(* Logix 5000 project; controller NWGG_Treater_Dayton vendor 1 type 14 code 238 rev 35.11; software revision 35.00 *)
// Treater at the Walla Walla Seed Plant

TASK MainTask (continuous, watchdog 500 ms) : MainProgram, Pumps, ColorBlending
TASK SafetyTask (periodic, rate 20 ms, priority 10, watchdog 20 ms, safety) : SafetyProgram

MODULES
   Local : vendor 1 type 14 code 238 (5069 0, rev 35.11)
      Pump_8 : PowerFlex 525-EENET (Ethernet 192.168.1.64, rev 7.1, Output RPI 20 ms)
      Pump_9 : PowerFlex 525-EENET (Ethernet 192.168.1.65, rev 7.1, Output RPI 20 ms)
      Pump_19 : PowerFlex 525-EENET (Ethernet 192.168.1.75, rev 7.1, Output RPI 20 ms)
      Pump_10 : PowerFlex 525-EENET (Ethernet 192.168.1.66, rev 7.1, Output RPI 20 ms)
      Pump_18 : PowerFlex 525-EENET (Ethernet 192.168.1.74, rev 7.1, Output RPI 20 ms)
      Pump_16 : PowerFlex 525-EENET (Ethernet 192.168.1.72, rev 7.1, Output RPI 20 ms)
      Pump_3 : PowerFlex 525-EENET (Ethernet 192.168.1.59, rev 7.1, Output RPI 20 ms)
      Treater_Drive : PowerFlex 525-EENET (Ethernet 192.168.1.81, rev 7.1, Output RPI 20 ms)
      Pump_21 : PowerFlex 525-EENET (Ethernet 192.168.1.77, rev 7.1, Output RPI 20 ms)
      Pump_6 : PowerFlex 525-EENET (Ethernet 192.168.1.62, rev 7.1, Output RPI 20 ms)
      Pump_20 : PowerFlex 525-EENET (Ethernet 192.168.1.76, rev 7.1, Output RPI 20 ms)
      Pump_22 : PowerFlex 525-EENET (Ethernet 192.168.1.78, rev 7.1, Output RPI 20 ms)
      Pump_14 : PowerFlex 525-EENET (Ethernet 192.168.1.70, rev 7.1, Output RPI 20 ms)
      Pump_13 : PowerFlex 525-EENET (Ethernet 192.168.1.69, rev 7.1, Output RPI 20 ms)
      Pump_15 : PowerFlex 525-EENET (Ethernet 192.168.1.71, rev 7.1, Output RPI 20 ms)
      Pump_7 : PowerFlex 525-EENET (Ethernet 192.168.1.63, rev 7.1, Output RPI 20 ms)
      Pump_5 : PowerFlex 525-EENET (Ethernet 192.168.1.61, rev 7.1, Output RPI 20 ms)
      Pump_12 : PowerFlex 525-EENET (Ethernet 192.168.1.68, rev 7.1, Output RPI 20 ms)
      Pump_2 : PowerFlex 525-EENET (Ethernet 192.168.1.58, rev 7.1, Output RPI 20 ms)
      Pump_1 : PowerFlex 525-EENET (Ethernet 192.168.1.57, rev 7.1, Output RPI 20 ms)
      Pump_11 : PowerFlex 525-EENET (Ethernet 192.168.1.67, rev 7.1, Output RPI 20 ms)
      Pump_17 : PowerFlex 525-EENET (Ethernet 192.168.1.73, rev 7.1, Output RPI 20 ms)
      Pump_4 : PowerFlex 525-EENET (Ethernet 192.168.1.60, rev 7.1, Output RPI 20 ms)
      Flex_IO_Adapter : 1794-AENTR (Ethernet 192.168.1.100, rev 1.1, Output RPI 20 ms)
         AC_Input : 1794-IA16 (Flex 2, rev 1.1)
         AC_Output : vendor 1 type 7 code 48 (Flex 3, rev 1.1)
         Analog_In_1 : vendor 1 type 10 code 25 (Flex 0, rev 2.1, Input RPI 80 ms)
         Analog_In_2 : vendor 1 type 10 code 25 (Flex 1, rev 2.1, Input RPI 80 ms)
      Scale_13 : vendor 666 type 12 code 16898 (Ethernet 192.168.1.123, rev 1.1, StandardDataDriven RPI 2 ms)
      Scale_22 : vendor 666 type 12 code 16898 (Ethernet 192.168.1.132, rev 1.1, StandardDataDriven RPI 2 ms)   // Pea Slurry
      Scale_9 : vendor 666 type 12 code 16898 (Ethernet 192.168.1.119, rev 1.1, StandardDataDriven RPI 2 ms)
      Scale_17 : vendor 666 type 12 code 16898 (Ethernet 192.168.1.127, rev 1.1, StandardDataDriven RPI 2 ms)
      Scale_8 : vendor 666 type 12 code 16898 (Ethernet 192.168.1.118, rev 1.1, StandardDataDriven RPI 2 ms)
      Scale_20 : vendor 666 type 12 code 16898 (Ethernet 192.168.1.130, rev 1.1, StandardDataDriven RPI 2 ms)
      Scale_19 : vendor 666 type 12 code 16898 (Ethernet 192.168.1.129, rev 1.1, StandardDataDriven RPI 2 ms)
      Scale_14 : vendor 666 type 12 code 16898 (Ethernet 192.168.1.124, rev 1.1, StandardDataDriven RPI 2 ms)
      Scale_6 : vendor 666 type 12 code 16898 (Ethernet 192.168.1.116, rev 1.1, StandardDataDriven RPI 2 ms)
      Scale_11 : vendor 666 type 12 code 16898 (Ethernet 192.168.1.121, rev 1.1, StandardDataDriven RPI 2 ms)
      Scale_21 : vendor 666 type 12 code 16898 (Ethernet 192.168.1.131, rev 1.1, StandardDataDriven RPI 2 ms)   // Small 3' By 3' Floor Scale
      Scale_1 : vendor 666 type 12 code 16898 (Ethernet 192.168.1.111, rev 1.1, StandardDataDriven RPI 2 ms)
      Scale_4 : vendor 666 type 12 code 16898 (Ethernet 192.168.1.114, rev 1.1, StandardDataDriven RPI 2 ms)
      Scale_18 : vendor 666 type 12 code 16898 (Ethernet 192.168.1.128, rev 1.1, StandardDataDriven RPI 2 ms)
      Scale_3 : vendor 666 type 12 code 16898 (Ethernet 192.168.1.113, rev 1.1, StandardDataDriven RPI 2 ms)
      Scale_5 : vendor 666 type 12 code 16898 (Ethernet 192.168.1.115, rev 1.1, StandardDataDriven RPI 2 ms)
      Scale_16 : vendor 666 type 12 code 16898 (Ethernet 192.168.1.126, rev 1.1, StandardDataDriven RPI 2 ms)
      Scale_2 : vendor 666 type 12 code 16898 (Ethernet 192.168.1.112, rev 1.1, StandardDataDriven RPI 2 ms)
      Scale_15 : vendor 666 type 12 code 16898 (Ethernet 192.168.1.125, rev 1.1, StandardDataDriven RPI 2 ms)
      Scale_10 : vendor 666 type 12 code 16898 (Ethernet 192.168.1.120, rev 1.1, StandardDataDriven RPI 2 ms)
      Scale_7 : vendor 666 type 12 code 16898 (Ethernet 192.168.1.117, rev 1.1, StandardDataDriven RPI 2 ms)
      Scale_12 : vendor 666 type 12 code 16898 (Ethernet 192.168.1.122, rev 1.1, StandardDataDriven RPI 2 ms)
      Water_Input : vendor 1 type 115 code 314 (5069 1, rev 2.1, StandardDataDriven RPI 100 ms)   // Input for Water Flow
END_MODULES

ADD_ON_INSTRUCTION Analog_Pump_Control   (* revision 1.0 *)
VAR_IN_OUT
   Pump_Drive_Out : AB:PowerFlex525V_EENET_Drive:O:0; {required}   // Pump Output
   Pump_Drive_In : AB:PowerFlex525V_EENET_Drive:I:0; {required}   // Pump Input
   Treater_Pump : Treater_Pump; {required}
        .Current_Oz_Rate   // This is the rate adjusted for the Current flow of grain reflected by the muiltliplier
END_VAR
VAR_INPUT
   Grain_Flow_CWT : REAL; {access None, required}
   Pump_Reversed : BOOL; {access Read Only, required}
END_VAR
VAR_IN_OUT
   Values : Analog_Gallon_Values; {required}   // Stored Values
   Analog_Raw_Counts : REAL; {required}
END_VAR
VAR_INPUT
   Start_Treating : BOOL; {access Read Only, required}
END_VAR
VAR
   Empty_String : STRING; {access None}
   PMC : Pump_Motor_Control; {access None}
   AnalogRate : Analog_Rate; {access None}
END_VAR

ROUTINE Logic   (* ladder *)
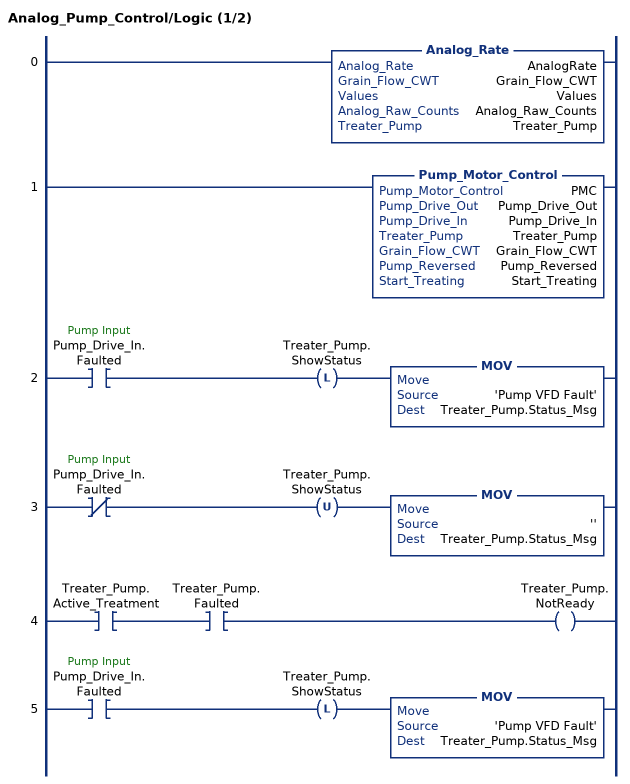
   0: Analog_Rate(AnalogRate,Grain_Flow_CWT,Values,Analog_Raw_Counts,Treater_Pump);
   1: Pump_Motor_Control(PMC,Pump_Drive_Out,Pump_Drive_In,Treater_Pump,Grain_Flow_CWT,Pump_Reversed,Start_Treating);
   2: XIC(Pump_Drive_In.Faulted)OTL(Treater_Pump.ShowStatus)MOV('Pump VFD Fault',Treater_Pump.Status_Msg);
   3: XIO(Pump_Drive_In.Faulted)OTU(Treater_Pump.ShowStatus)MOV('',Treater_Pump.Status_Msg);
   4: XIC(Treater_Pump.Active_Treatment)XIC(Treater_Pump.Faulted)OTE(Treater_Pump.NotReady);
   5: XIC(Pump_Drive_In.Faulted)OTL(Treater_Pump.ShowStatus)MOV('Pump VFD Fault',Treater_Pump.Status_Msg);
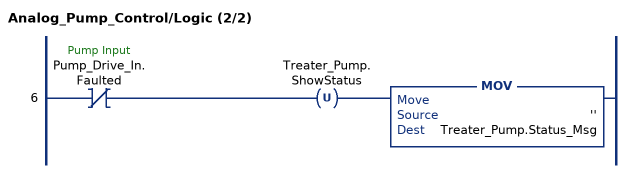
   6: XIO(Pump_Drive_In.Faulted)OTU(Treater_Pump.ShowStatus)MOV('',Treater_Pump.Status_Msg);
END_ROUTINE
END_ADD_ON_INSTRUCTION

ADD_ON_INSTRUCTION Analog_Rate   (* revision 1.0 *)
VAR_INPUT
   Grain_Flow_CWT : REAL; {access None, required}
END_VAR
VAR_IN_OUT
   Values : Analog_Gallon_Values; {required}   // Stored Values
END_VAR
VAR_INPUT
   Analog_Raw_Counts : REAL; {access Read Only, required}   // Values From CT
END_VAR
VAR_IN_OUT
   Treater_Pump : Treater_Pump; {required}
END_VAR

ROUTINE Logic   (* ladder *)
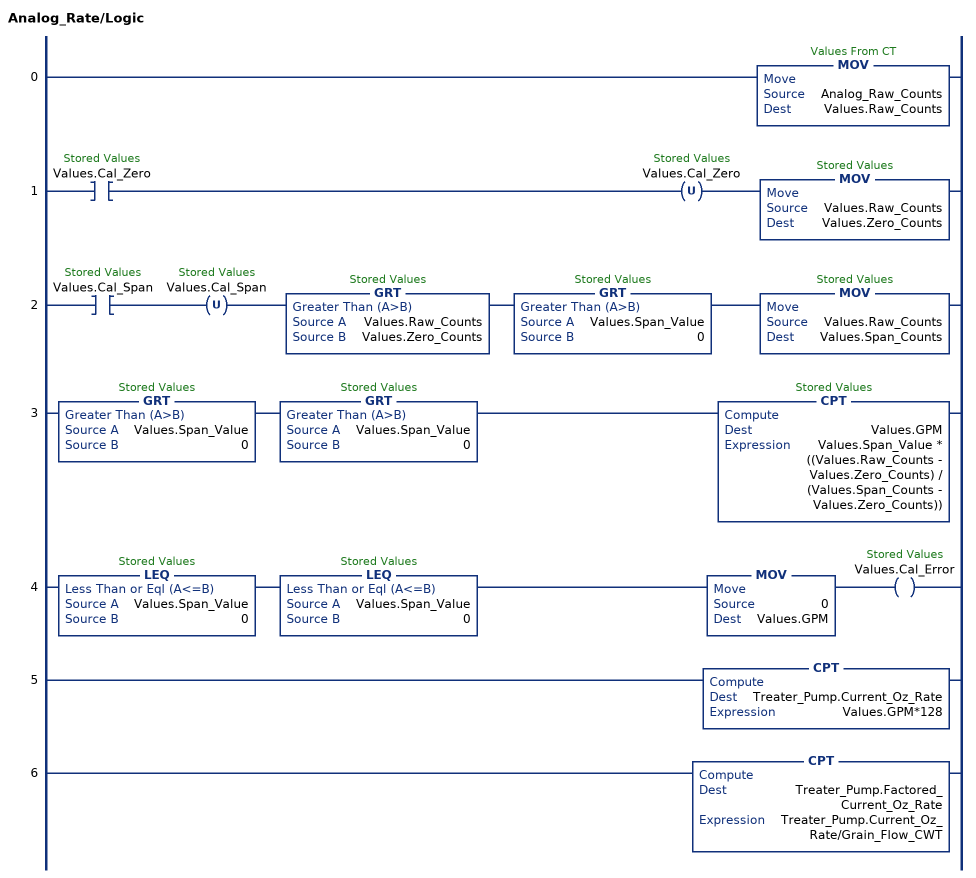
   0: MOV(Analog_Raw_Counts,Values.Raw_Counts);
   1: XIC(Values.Cal_Zero)OTU(Values.Cal_Zero)MOV(Values.Raw_Counts,Values.Zero_Counts);
   2: XIC(Values.Cal_Span)OTU(Values.Cal_Span)GRT(Values.Raw_Counts,Values.Zero_Counts)GRT(Values.Span_Value,0)MOV(Values.Raw_Counts,Values.Span_Counts);
   3: GRT(Values.Span_Value,0)GRT(Values.Span_Value,0)CPT(Values.GPM,Values.Span_Value * ((Values.Raw_Counts - Values.Zero_Counts) / (Values.Span_Counts - Values.Zero_Counts)));
   4: LEQ(Values.Span_Value,0)LEQ(Values.Span_Value,0)MOV(0,Values.GPM)OTE(Values.Cal_Error);
   5: CPT(Treater_Pump.Current_Oz_Rate,Values.GPM*128);
   6: CPT(Treater_Pump.Factored_Current_Oz_Rate,Treater_Pump.Current_Oz_Rate/Grain_Flow_CWT);
END_ROUTINE
END_ADD_ON_INSTRUCTION

ADD_ON_INSTRUCTION ColorBlending   (* revision 1.0 *)
VAR_IN_OUT
   White_Pump : Treater_Pump; {required}
   Blue_Pump : Treater_Pump; {required}
   Yellow_Pump : Treater_Pump; {required}
   Red_Pump : Treater_Pump; {required}
   Polymer_Pump : Treater_Pump; {required}
   SelectedColors : Color[10]; {required}
END_VAR
VAR_INPUT
   Reset : BOOL;
   Start : BOOL;
   Total_Oz_Min : REAL; {access None}
   PumpDelay : DINT;
   ReverseDuration : DINT;
   Pause : BOOL;
END_VAR
VAR
   Current_Color_Index : COUNTER; {access Read Only}
   tmrDuration : TIMER; {access None}
   Current_Color : Color; {access None}
   tmrDelay : TIMER; {access None}
   tmrReverse : TIMER; {access None}
   Inactive_Color : BOOL; {access None}
END_VAR

ROUTINE Logic   (* ladder *)
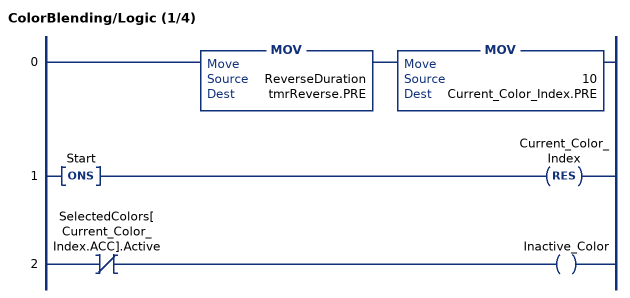
   0: MOV(ReverseDuration,tmrReverse.PRE)MOV(10,Current_Color_Index.PRE);
   1: ONS(Start)RES(Current_Color_Index);
   2: XIO(SelectedColors[Current_Color_Index.ACC].Active)OTE(Inactive_Color);
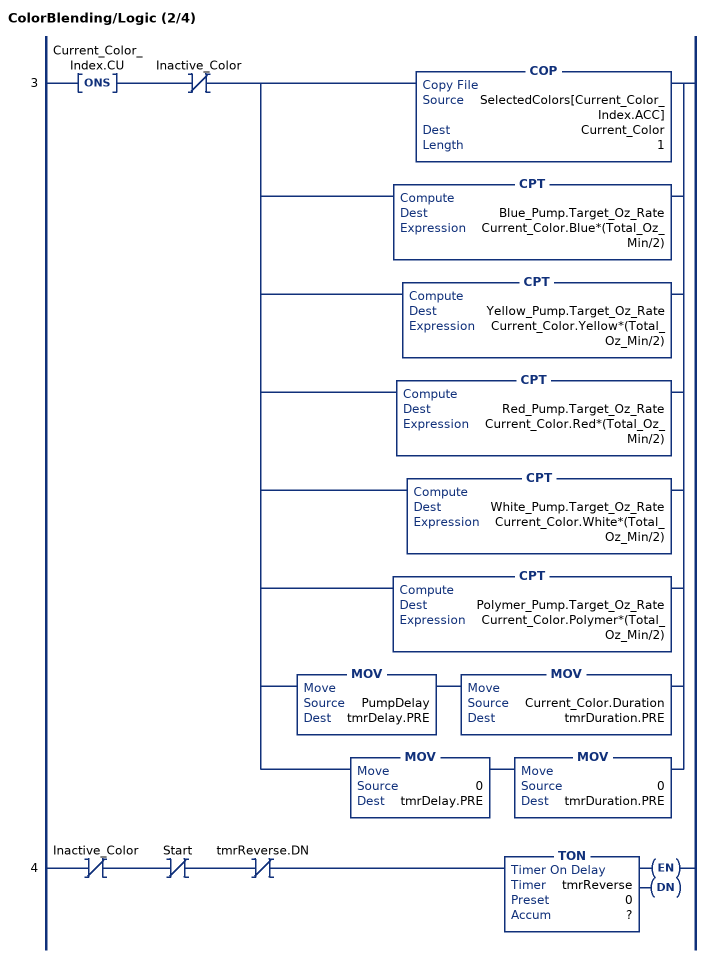
   3: ONS(Current_Color_Index.CU)XIO(Inactive_Color)[COP(SelectedColors[Current_Color_Index.ACC],Current_Color,1) ,CPT(Blue_Pump.Target_Oz_Rate,Current_Color.Blue*(Total_Oz_Min/2)) ,CPT(Yellow_Pump.Target_Oz_Rate,Current_Color.Yellow*(Total_Oz_Min/2)) ,CPT(Red_Pump.Target_Oz_Rate,Current_Color.Red*(Total_Oz_Min/2)) ,CPT(White_Pump.Target_Oz_Rate,Current_Color.White*(Total_Oz_Min/2)) ,CPT(Polymer_Pump.Target_Oz_Rate,Current_Color.Polymer*(Total_Oz_Min/2)) ,MOV(PumpDelay,tmrDelay.PRE) MOV(Current_Color.Duration,tmrDuration.PRE) ,MOV(0,tmrDelay.PRE) MOV(0,tmrDuration.PRE) ];
   4: XIO(Inactive_Color)XIO(Start)XIO(tmrReverse.DN)TON(tmrReverse,?,?);
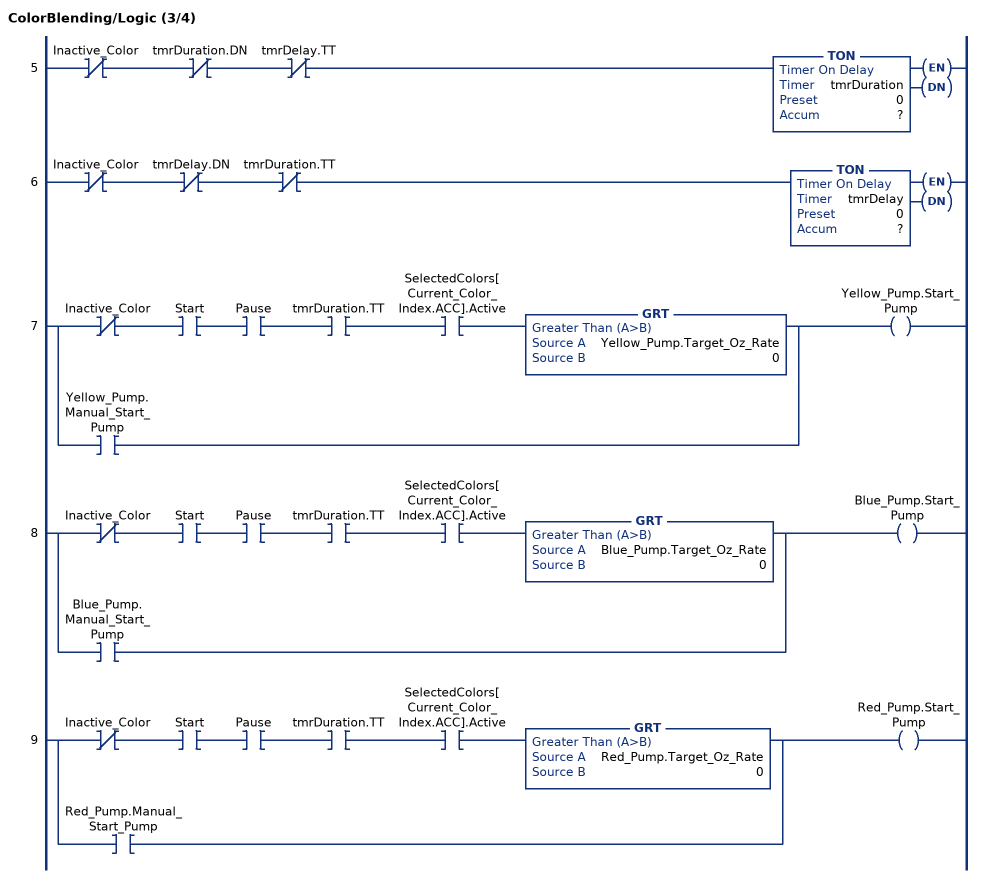
   5: XIO(Inactive_Color)XIO(tmrDuration.DN)XIO(tmrDelay.TT)TON(tmrDuration,?,?);
   6: XIO(Inactive_Color)XIO(tmrDelay.DN)XIO(tmrDuration.TT)TON(tmrDelay,?,?);
   7: [XIO(Inactive_Color) XIC(Start) XIC(Pause) XIC(tmrDuration.TT) XIC(SelectedColors[Current_Color_Index.ACC].Active) GRT(Yellow_Pump.Target_Oz_Rate,0) ,XIC(Yellow_Pump.Manual_Start_Pump) ]OTE(Yellow_Pump.Start_Pump);
   8: [XIO(Inactive_Color) XIC(Start) XIC(Pause) XIC(tmrDuration.TT) XIC(SelectedColors[Current_Color_Index.ACC].Active) GRT(Blue_Pump.Target_Oz_Rate,0) ,XIC(Blue_Pump.Manual_Start_Pump) ]OTE(Blue_Pump.Start_Pump);
   9: [XIO(Inactive_Color) XIC(Start) XIC(Pause) XIC(tmrDuration.TT) XIC(SelectedColors[Current_Color_Index.ACC].Active) GRT(Red_Pump.Target_Oz_Rate,0) ,XIC(Red_Pump.Manual_Start_Pump) ]OTE(Red_Pump.Start_Pump);
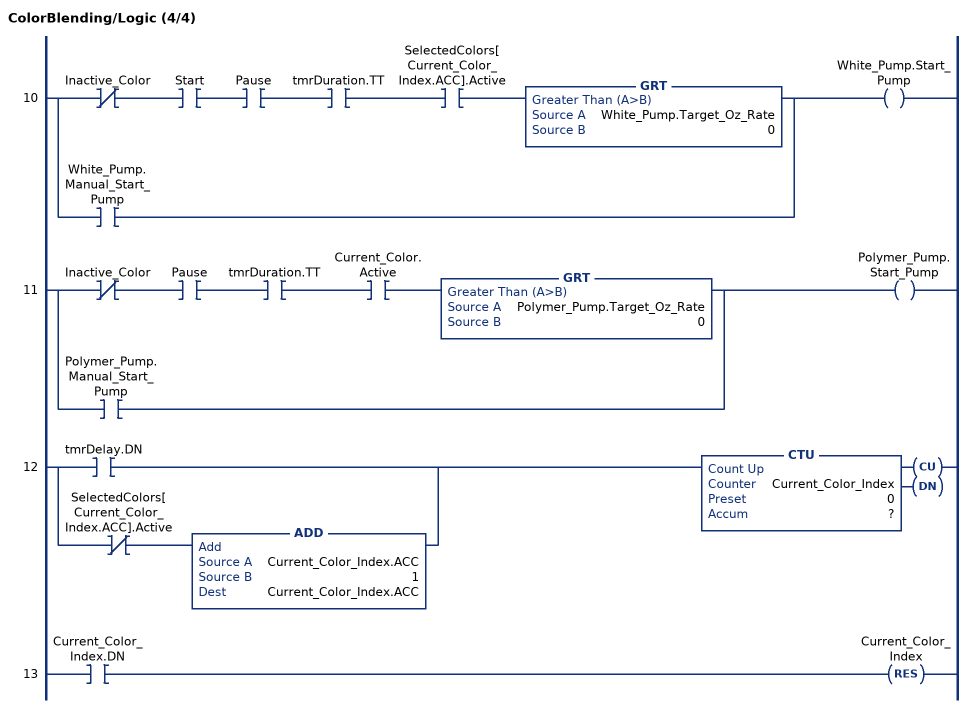
   10: [XIO(Inactive_Color) XIC(Start) XIC(Pause) XIC(tmrDuration.TT) XIC(SelectedColors[Current_Color_Index.ACC].Active) GRT(White_Pump.Target_Oz_Rate,0) ,XIC(White_Pump.Manual_Start_Pump) ]OTE(White_Pump.Start_Pump);
   11: [XIO(Inactive_Color) XIC(Pause) XIC(tmrDuration.TT) XIC(Current_Color.Active) GRT(Polymer_Pump.Target_Oz_Rate,0) ,XIC(Polymer_Pump.Manual_Start_Pump) ]OTE(Polymer_Pump.Start_Pump);
   12: [XIC(tmrDelay.DN) ,XIO(SelectedColors[Current_Color_Index.ACC].Active) ADD(Current_Color_Index.ACC,1,Current_Color_Index.ACC) ]CTU(Current_Color_Index,?,?);
   13: XIC(Current_Color_Index.DN)RES(Current_Color_Index);
END_ROUTINE
END_ADD_ON_INSTRUCTION

ADD_ON_INSTRUCTION Get_Active_Pumps   (* revision 1.0 *)
VAR_IN_OUT
   Treater_Pump : Treater_Pump[50]; {required}
   Active_Pump : Active_Pump_Values[10]; {required}
END_VAR
VAR
   Active_Pump_Count : DINT; {access None}
END_VAR

ROUTINE Logic   (* ladder *)
END_ROUTINE
END_ADD_ON_INSTRUCTION

ADD_ON_INSTRUCTION Pump_Motor_Control   (* revision 1.0 *)
VAR_IN_OUT
   Pump_Drive_Out : AB:PowerFlex525V_EENET_Drive:O:0; {required}   // Pump Output
   Pump_Drive_In : AB:PowerFlex525V_EENET_Drive:I:0; {required}   // Pump Input
   Treater_Pump : Treater_Pump; {required}
        .Current_Oz_Rate   // This is the rate adjusted for the Current flow of grain reflected by the muiltliplier
END_VAR
VAR_INPUT
   Grain_Flow_CWT : REAL; {access None, required}
   Pump_Reversed : BOOL; {access Read Only, required}
   Start_Treating : BOOL; {access Read Only, required}
END_VAR
VAR
   OverSpeedLimit : DINT; {access None}
   tmrOverSpeed : TIMER; {access None}
   PumpTreatingOn : BOOL; {access None}
   tmrPIDDelay : TIMER; {access None}
   tmrOverSpeedReset : TIMER; {access None}
   Reset_New_Product : BOOL; {access None}
   Empty_String : STRING; {access None}
END_VAR

ROUTINE Logic   (* ladder *)
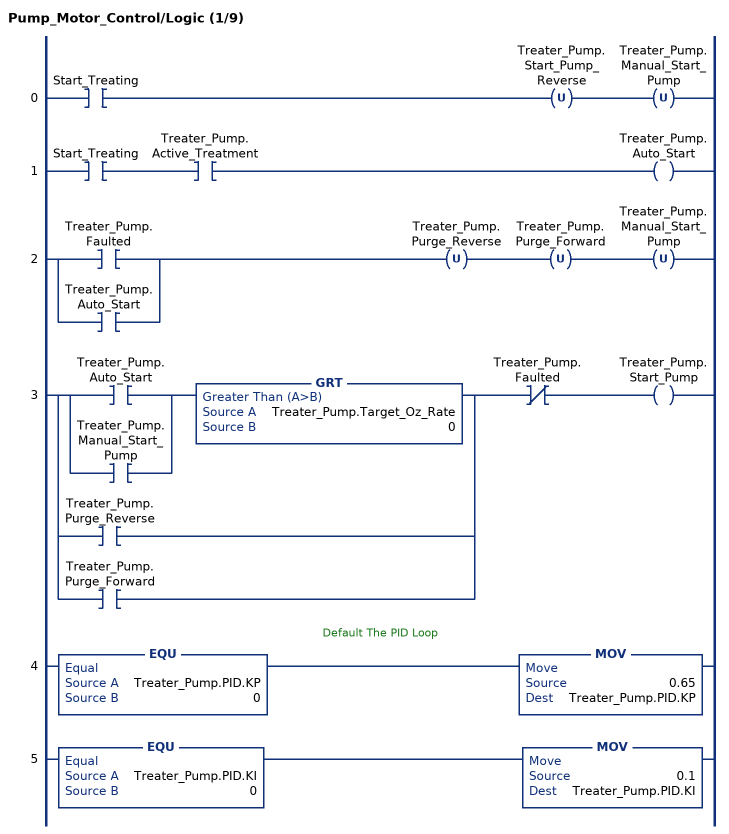
   0: XIC(Start_Treating)OTU(Treater_Pump.Start_Pump_Reverse)OTU(Treater_Pump.Manual_Start_Pump);
   1: XIC(Start_Treating)XIC(Treater_Pump.Active_Treatment)OTE(Treater_Pump.Auto_Start);
   2: [XIC(Treater_Pump.Faulted) ,XIC(Treater_Pump.Auto_Start) ]OTU(Treater_Pump.Purge_Reverse)OTU(Treater_Pump.Purge_Forward)OTU(Treater_Pump.Manual_Start_Pump);
   3: [[XIC(Treater_Pump.Auto_Start) ,XIC(Treater_Pump.Manual_Start_Pump) ] GRT(Treater_Pump.Target_Oz_Rate,0) ,XIC(Treater_Pump.Purge_Reverse) ,XIC(Treater_Pump.Purge_Forward) ]XIO(Treater_Pump.Faulted)OTE(Treater_Pump.Start_Pump);
   // Default The PID Loop
   4: EQU(Treater_Pump.PID.KP,0)MOV(0.65,Treater_Pump.PID.KP);
   5: EQU(Treater_Pump.PID.KI,0)MOV(0.1,Treater_Pump.PID.KI);
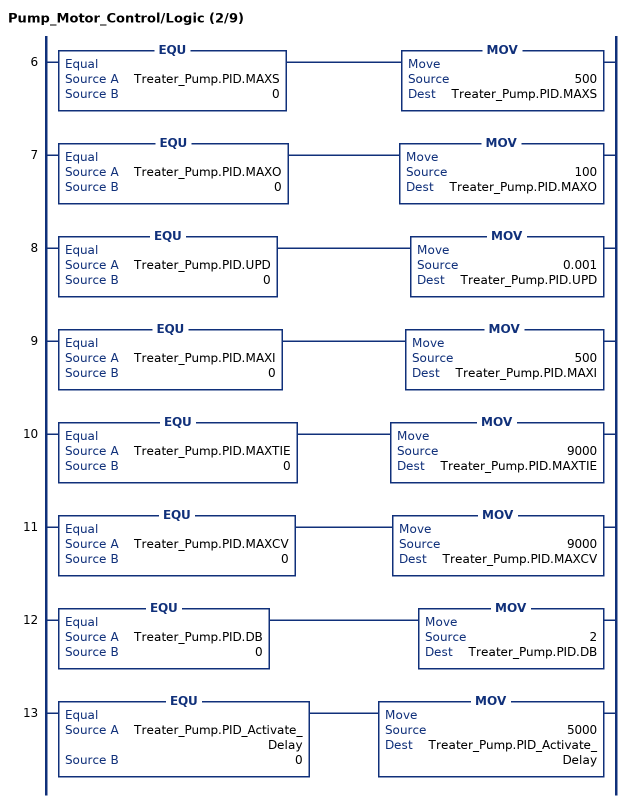
   6: EQU(Treater_Pump.PID.MAXS,0)MOV(500,Treater_Pump.PID.MAXS);
   7: EQU(Treater_Pump.PID.MAXO,0)MOV(100,Treater_Pump.PID.MAXO);
   8: EQU(Treater_Pump.PID.UPD,0)MOV(0.001,Treater_Pump.PID.UPD);
   9: EQU(Treater_Pump.PID.MAXI,0)MOV(500,Treater_Pump.PID.MAXI);
   10: EQU(Treater_Pump.PID.MAXTIE,0)MOV(9000,Treater_Pump.PID.MAXTIE);
   11: EQU(Treater_Pump.PID.MAXCV,0)MOV(9000,Treater_Pump.PID.MAXCV);
   12: EQU(Treater_Pump.PID.DB,0)MOV(2,Treater_Pump.PID.DB);
   13: EQU(Treater_Pump.PID_Activate_Delay,0)MOV(5000,Treater_Pump.PID_Activate_Delay);
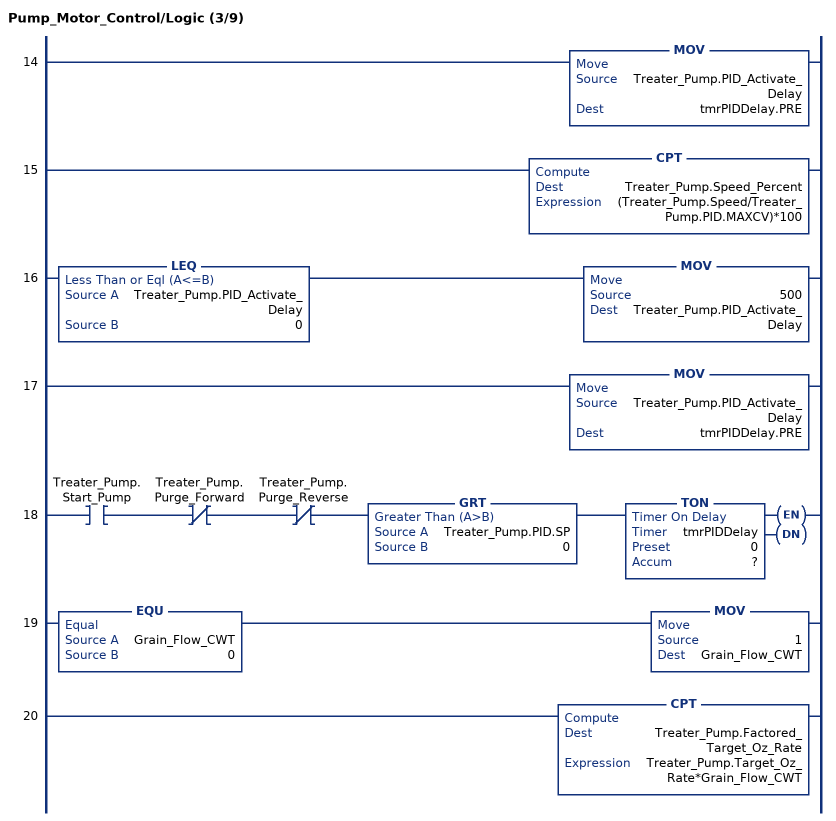
   14: MOV(Treater_Pump.PID_Activate_Delay,tmrPIDDelay.PRE);
   15: CPT(Treater_Pump.Speed_Percent,(Treater_Pump.Speed/Treater_Pump.PID.MAXCV)*100);
   16: LEQ(Treater_Pump.PID_Activate_Delay,0)MOV(500,Treater_Pump.PID_Activate_Delay);
   17: MOV(Treater_Pump.PID_Activate_Delay,tmrPIDDelay.PRE);
   18: XIC(Treater_Pump.Start_Pump)XIO(Treater_Pump.Purge_Forward)XIO(Treater_Pump.Purge_Reverse)GRT(Treater_Pump.PID.SP,0)TON(tmrPIDDelay,?,?);
   19: EQU(Grain_Flow_CWT,0)MOV(1,Grain_Flow_CWT);
   20: CPT(Treater_Pump.Factored_Target_Oz_Rate,Treater_Pump.Target_Oz_Rate*Grain_Flow_CWT);
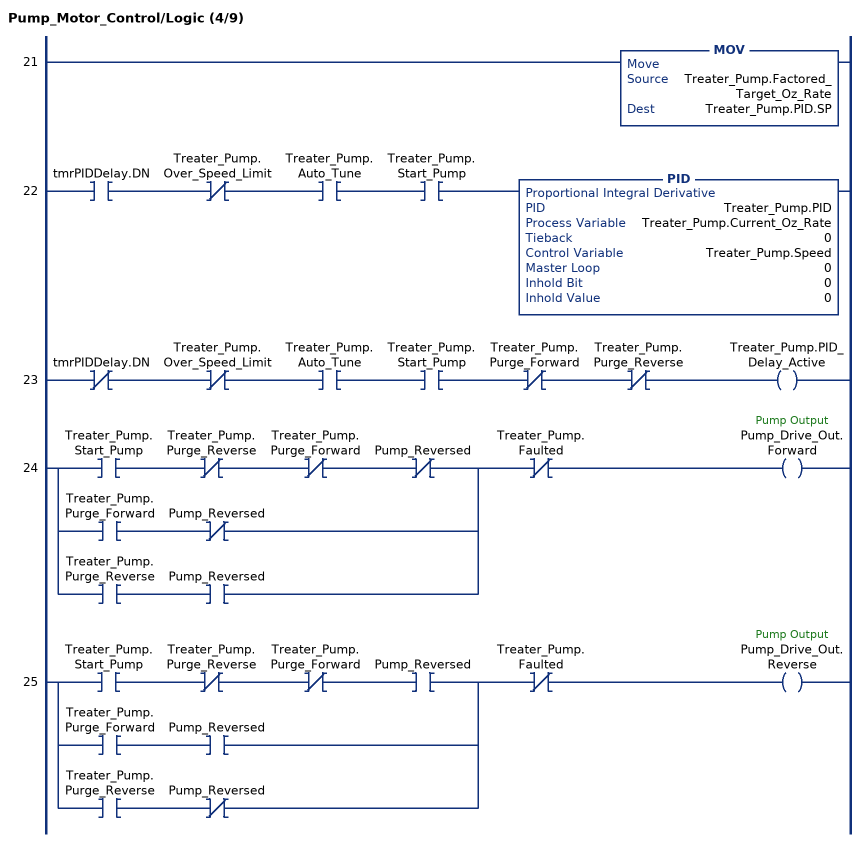
   21: MOV(Treater_Pump.Factored_Target_Oz_Rate,Treater_Pump.PID.SP);
   22: XIC(tmrPIDDelay.DN)XIO(Treater_Pump.Over_Speed_Limit)XIC(Treater_Pump.Auto_Tune)XIC(Treater_Pump.Start_Pump)PID(Treater_Pump.PID,Treater_Pump.Current_Oz_Rate,0,Treater_Pump.Speed,0,0,0);
   23: XIO(tmrPIDDelay.DN)XIO(Treater_Pump.Over_Speed_Limit)XIC(Treater_Pump.Auto_Tune)XIC(Treater_Pump.Start_Pump)XIO(Treater_Pump.Purge_Forward)XIO(Treater_Pump.Purge_Reverse)OTE(Treater_Pump.PID_Delay_Active);
   24: [XIC(Treater_Pump.Start_Pump) XIO(Treater_Pump.Purge_Reverse) XIO(Treater_Pump.Purge_Forward) XIO(Pump_Reversed) ,XIC(Treater_Pump.Purge_Forward) XIO(Pump_Reversed) ,XIC(Treater_Pump.Purge_Reverse) XIC(Pump_Reversed) ]XIO(Treater_Pump.Faulted)OTE(Pump_Drive_Out.Forward);
   25: [XIC(Treater_Pump.Start_Pump) XIO(Treater_Pump.Purge_Reverse) XIO(Treater_Pump.Purge_Forward) XIC(Pump_Reversed) ,XIC(Treater_Pump.Purge_Forward) XIC(Pump_Reversed) ,XIC(Treater_Pump.Purge_Reverse) XIO(Pump_Reversed) ]XIO(Treater_Pump.Faulted)OTE(Pump_Drive_Out.Reverse);
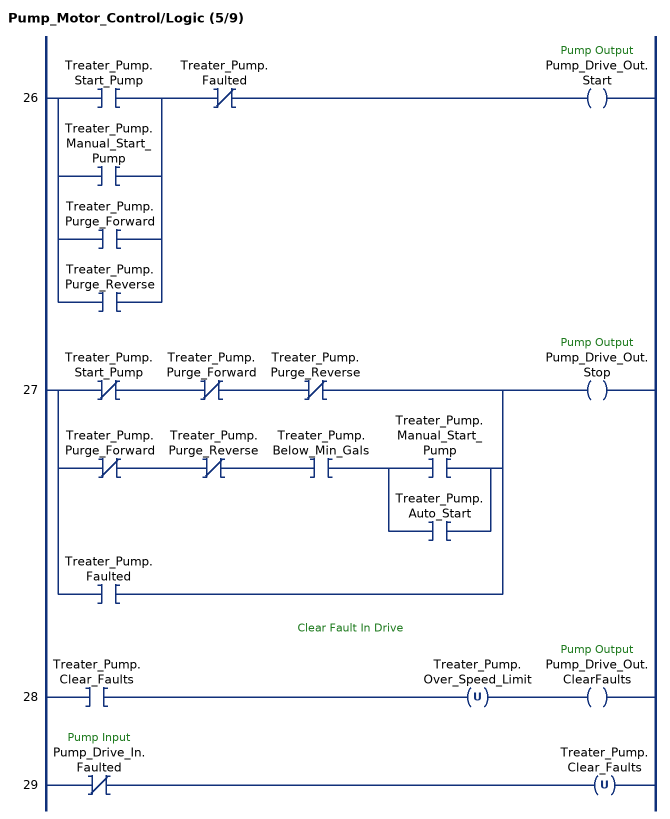
   26: [XIC(Treater_Pump.Start_Pump) ,XIC(Treater_Pump.Manual_Start_Pump) ,XIC(Treater_Pump.Purge_Forward) ,XIC(Treater_Pump.Purge_Reverse) ]XIO(Treater_Pump.Faulted)OTE(Pump_Drive_Out.Start);
   27: [XIO(Treater_Pump.Start_Pump) XIO(Treater_Pump.Purge_Forward) XIO(Treater_Pump.Purge_Reverse) ,XIO(Treater_Pump.Purge_Forward) XIO(Treater_Pump.Purge_Reverse) XIC(Treater_Pump.Below_Min_Gals) [XIC(Treater_Pump.Manual_Start_Pump) ,XIC(Treater_Pump.Auto_Start) ] ,XIC(Treater_Pump.Faulted) ]OTE(Pump_Drive_Out.Stop);
   // Clear Fault In Drive
   28: XIC(Treater_Pump.Clear_Faults)OTU(Treater_Pump.Over_Speed_Limit)OTE(Pump_Drive_Out.ClearFaults);
   29: XIO(Pump_Drive_In.Faulted)OTU(Treater_Pump.Clear_Faults);
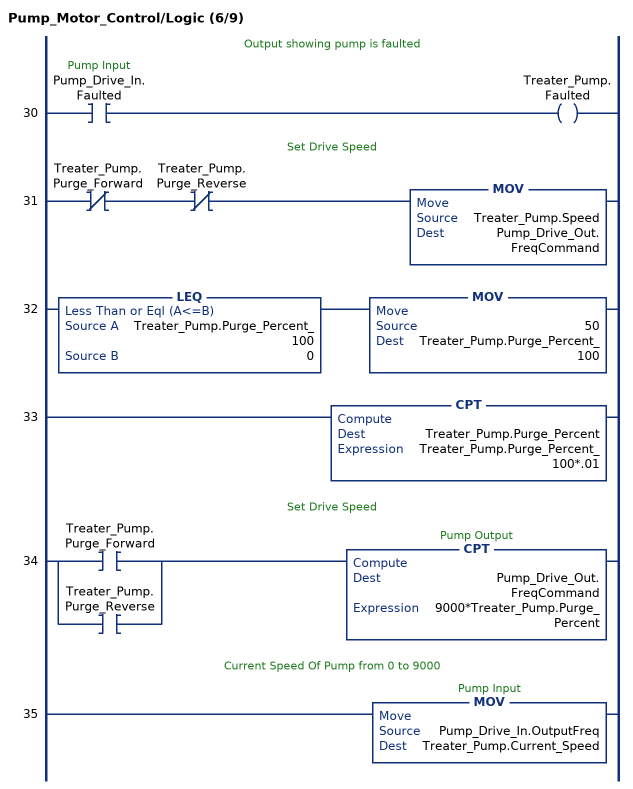
   // Output showing pump is faulted
   30: XIC(Pump_Drive_In.Faulted)OTE(Treater_Pump.Faulted);
   // Set Drive Speed
   31: XIO(Treater_Pump.Purge_Forward)XIO(Treater_Pump.Purge_Reverse)MOV(Treater_Pump.Speed,Pump_Drive_Out.FreqCommand);
   32: LEQ(Treater_Pump.Purge_Percent_100,0)MOV(50,Treater_Pump.Purge_Percent_100);
   33: CPT(Treater_Pump.Purge_Percent,Treater_Pump.Purge_Percent_100*.01);
   // Set Drive Speed
   34: [XIC(Treater_Pump.Purge_Forward) ,XIC(Treater_Pump.Purge_Reverse) ]CPT(Pump_Drive_Out.FreqCommand,9000*Treater_Pump.Purge_Percent);
   // Current Speed Of Pump from 0 to 9000
   35: MOV(Pump_Drive_In.OutputFreq,Treater_Pump.Current_Speed);
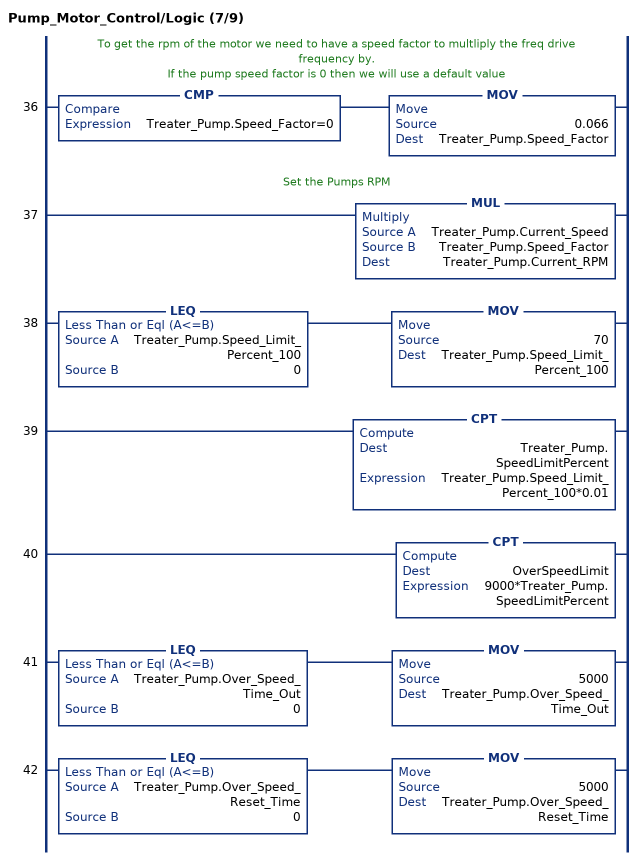
   // To get the rpm of the motor we need to have a speed factor to multliply the freq drive frequency by.
   // If the pump speed factor is 0 then we will use a default value
   36: CMP(Treater_Pump.Speed_Factor=0)MOV(0.066,Treater_Pump.Speed_Factor);
   // Set the Pumps RPM
   37: MUL(Treater_Pump.Current_Speed,Treater_Pump.Speed_Factor,Treater_Pump.Current_RPM);
   38: LEQ(Treater_Pump.Speed_Limit_Percent_100,0)MOV(70,Treater_Pump.Speed_Limit_Percent_100);
   39: CPT(Treater_Pump.SpeedLimitPercent,Treater_Pump.Speed_Limit_Percent_100*0.01);
   40: CPT(OverSpeedLimit,9000*Treater_Pump.SpeedLimitPercent);
   41: LEQ(Treater_Pump.Over_Speed_Time_Out,0)MOV(5000,Treater_Pump.Over_Speed_Time_Out);
   42: LEQ(Treater_Pump.Over_Speed_Reset_Time,0)MOV(5000,Treater_Pump.Over_Speed_Reset_Time);
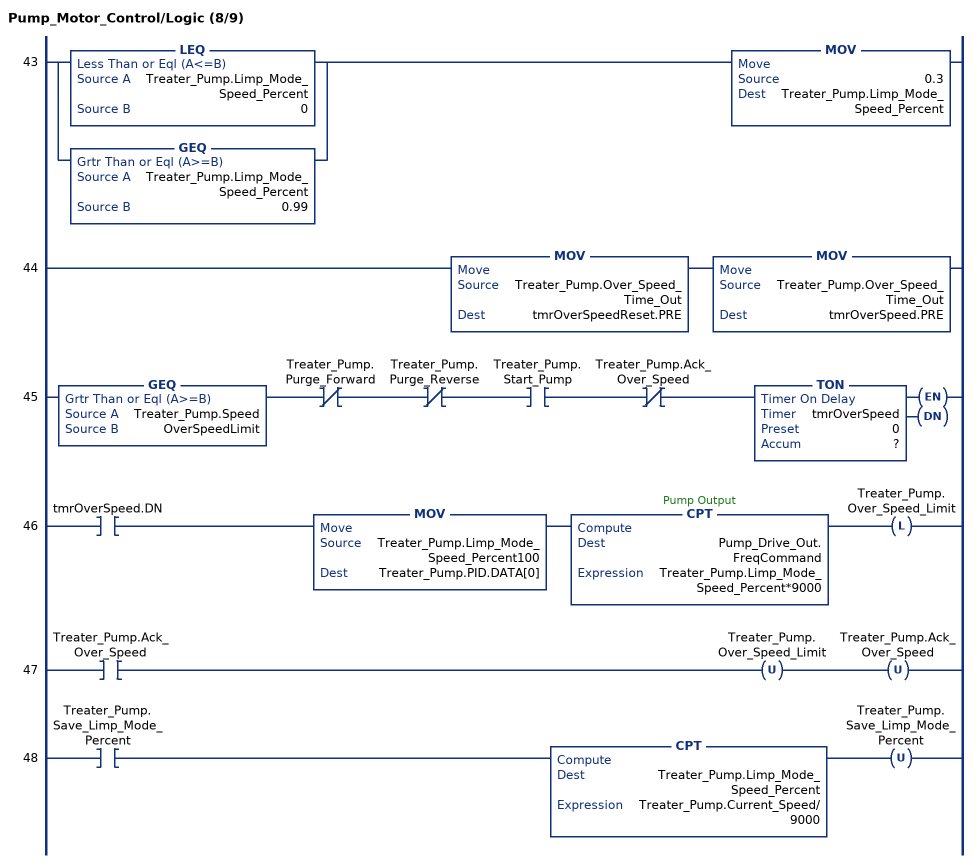
   43: [LEQ(Treater_Pump.Limp_Mode_Speed_Percent,0) ,GEQ(Treater_Pump.Limp_Mode_Speed_Percent,0.99) ]MOV(0.3,Treater_Pump.Limp_Mode_Speed_Percent);
   44: MOV(Treater_Pump.Over_Speed_Time_Out,tmrOverSpeedReset.PRE)MOV(Treater_Pump.Over_Speed_Time_Out,tmrOverSpeed.PRE);
   45: GEQ(Treater_Pump.Speed,OverSpeedLimit)XIO(Treater_Pump.Purge_Forward)XIO(Treater_Pump.Purge_Reverse)XIC(Treater_Pump.Start_Pump)XIO(Treater_Pump.Ack_Over_Speed)TON(tmrOverSpeed,?,?);
   46: XIC(tmrOverSpeed.DN)MOV(Treater_Pump.Limp_Mode_Speed_Percent100,Treater_Pump.PID.DATA[0])CPT(Pump_Drive_Out.FreqCommand,Treater_Pump.Limp_Mode_Speed_Percent*9000)OTL(Treater_Pump.Over_Speed_Limit);
   47: XIC(Treater_Pump.Ack_Over_Speed)OTU(Treater_Pump.Over_Speed_Limit)OTU(Treater_Pump.Ack_Over_Speed);
   48: XIC(Treater_Pump.Save_Limp_Mode_Percent)CPT(Treater_Pump.Limp_Mode_Speed_Percent,Treater_Pump.Current_Speed/9000)OTU(Treater_Pump.Save_Limp_Mode_Percent);
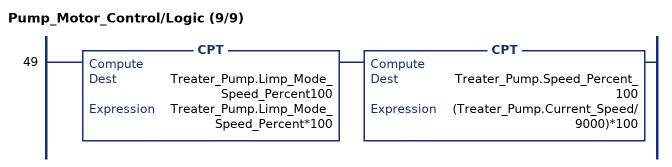
   49: CPT(Treater_Pump.Limp_Mode_Speed_Percent100,Treater_Pump.Limp_Mode_Speed_Percent*100)CPT(Treater_Pump.Speed_Percent_100,(Treater_Pump.Current_Speed/9000)*100);
END_ROUTINE
END_ADD_ON_INSTRUCTION

ADD_ON_INSTRUCTION Pump_Scale_Control   (* revision 1.0 *)
VAR_IN_OUT
   Pump_Drive_Out : AB:PowerFlex525V_EENET_Drive:O:0; {required}   // Pump Output
        .Reverse   // Pump is installed backwards So Reverse is forward
   Pump_Drive_In : AB:PowerFlex525V_EENET_Drive:I:0; {required}   // Pump Input
   Treater_Pump : Treater_Pump; {required}
END_VAR
VAR_INPUT
   Grain_Flow_CWT : REAL; {access None, required}
   Pump_Reversed : BOOL; {access Read Only, required}
   Start_Treating : BOOL; {access Read Only, required}
END_VAR
VAR
   SAIScaleRate : SAI_Scale_Rate; {access None}
   PMC : Pump_Motor_Control; {access None}
END_VAR

ROUTINE Logic   (* ladder *)
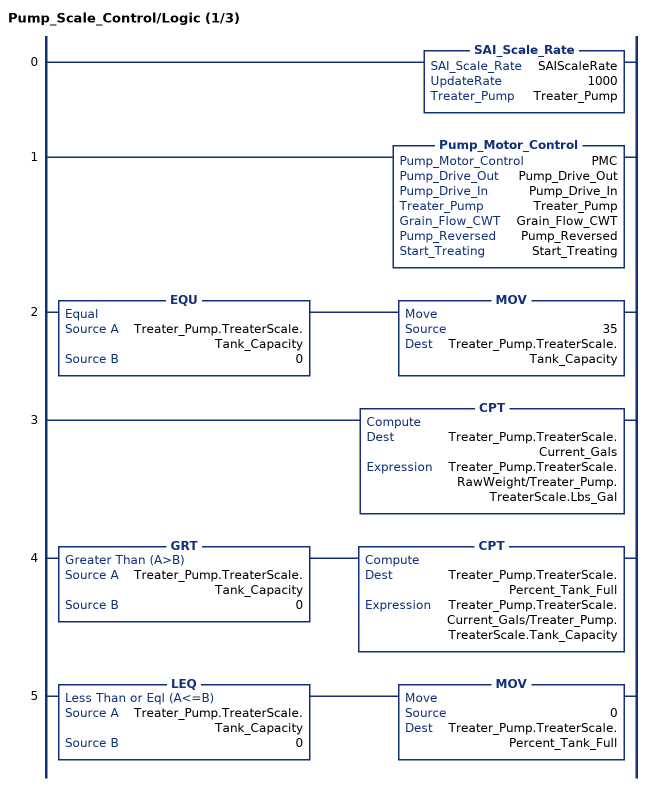
   0: SAI_Scale_Rate(SAIScaleRate,1000,Treater_Pump);
   1: Pump_Motor_Control(PMC,Pump_Drive_Out,Pump_Drive_In,Treater_Pump,Grain_Flow_CWT,Pump_Reversed,Start_Treating);
   2: EQU(Treater_Pump.TreaterScale.Tank_Capacity,0)MOV(35,Treater_Pump.TreaterScale.Tank_Capacity);
   3: CPT(Treater_Pump.TreaterScale.Current_Gals,Treater_Pump.TreaterScale.RawWeight/Treater_Pump.TreaterScale.Lbs_Gal);
   4: GRT(Treater_Pump.TreaterScale.Tank_Capacity,0)CPT(Treater_Pump.TreaterScale.Percent_Tank_Full,Treater_Pump.TreaterScale.Current_Gals/Treater_Pump.TreaterScale.Tank_Capacity);
   5: LEQ(Treater_Pump.TreaterScale.Tank_Capacity,0)MOV(0,Treater_Pump.TreaterScale.Percent_Tank_Full);
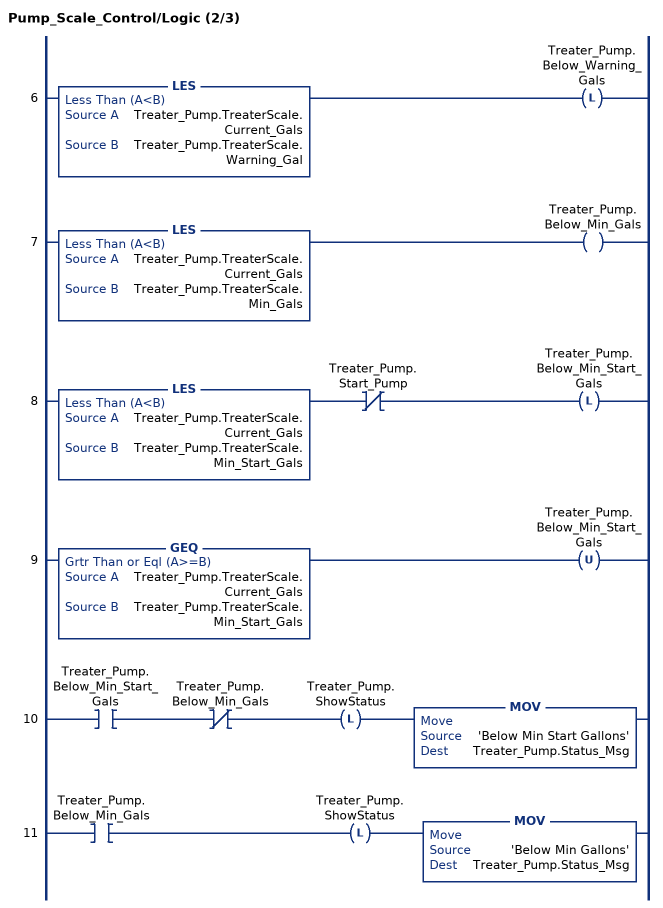
   6: LES(Treater_Pump.TreaterScale.Current_Gals,Treater_Pump.TreaterScale.Warning_Gal)OTL(Treater_Pump.Below_Warning_Gals);
   7: LES(Treater_Pump.TreaterScale.Current_Gals,Treater_Pump.TreaterScale.Min_Gals)OTE(Treater_Pump.Below_Min_Gals);
   8: LES(Treater_Pump.TreaterScale.Current_Gals,Treater_Pump.TreaterScale.Min_Start_Gals)XIO(Treater_Pump.Start_Pump)OTL(Treater_Pump.Below_Min_Start_Gals);
   9: GEQ(Treater_Pump.TreaterScale.Current_Gals,Treater_Pump.TreaterScale.Min_Start_Gals)OTU(Treater_Pump.Below_Min_Start_Gals);
   10: XIC(Treater_Pump.Below_Min_Start_Gals)XIO(Treater_Pump.Below_Min_Gals)OTL(Treater_Pump.ShowStatus)MOV('Below Min Start Gallons',Treater_Pump.Status_Msg);
   11: XIC(Treater_Pump.Below_Min_Gals)OTL(Treater_Pump.ShowStatus)MOV('Below Min Gallons',Treater_Pump.Status_Msg);
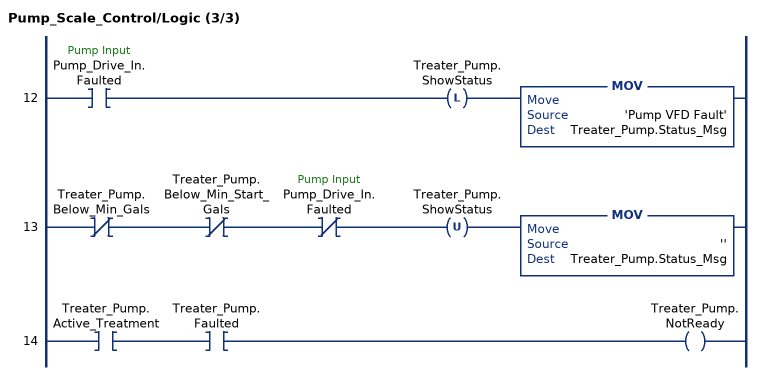
   12: XIC(Pump_Drive_In.Faulted)OTL(Treater_Pump.ShowStatus)MOV('Pump VFD Fault',Treater_Pump.Status_Msg);
   13: XIO(Treater_Pump.Below_Min_Gals)XIO(Treater_Pump.Below_Min_Start_Gals)XIO(Pump_Drive_In.Faulted)OTU(Treater_Pump.ShowStatus)MOV('',Treater_Pump.Status_Msg);
   14: XIC(Treater_Pump.Active_Treatment)XIC(Treater_Pump.Faulted)OTE(Treater_Pump.NotReady);
END_ROUTINE
END_ADD_ON_INSTRUCTION
